(* CODESYS project liang test485.project

Project tree, tasks and I/O mapping:
  Device : AM402-CPU1608TP/TN, Shenzhen Inovance Control Technology, version 3.5.11.11
    application Application
      libraries: Standard, * (System)
      task MainTask (cyclic, interval 4 ms, priority 1) calls PLC_PRG
      program PLC_PRG [ST]
      DifferentialMonitor
      data type ST_MBTask
      program FB_ModbusRTU_Poller [ST]
    HardWare Configuration
    Network Configuration
      LocalBus Config
    Device Diagnosis
    Resources List
    ConfigStorage
    SoftMotion General Axis Pool
    HIGH_SPEED_IO : 高速IO模块, Inovance, version 00.00.00.20
        unmapped channels: InputData, OutputData
      HSIO
    MODBUS_COM0 : Modbus主站, inovance, version 00.00.00.10
        settings: Vendor.parameterset.Bit0 = False; Vendor.res = 0;  = 0
      modbus_protocol : Modbus Slave, Inovance, version 00.00.00.10
          settings: UseDec = False; modbus slave com port.ChannelNum = 3; modbus slave com port.EnableSlaveVariable = 1001; channel.PremeterSet.Bit2 = TRUE; channel.PremeterSet.Bit4 = TRUE; channel.CycleTimes = 500; channel.ReadRegOffSet = 0; channel.WriteRegOffSet = 8193; channel.IOChannel = 0; channel.ResendCount = 1; channel.ChannelName = '写频率'; channel.ChannelNote = ''; channel.PremeterSet.Bit2 = TRUE; channel.PremeterSet.Bit4 = TRUE; channel.ReadRegOffSet = 0; channel.WriteRegOffSet = 8192; channel.ResendCount = 1; channel.ChannelName = '写控制字'; channel.ChannelNote = ''; channel.PremeterSet.Bit3 = TRUE; channel.ReadRegOffSet = 8448; channel.ReadRegLeg = 4; channel.WriteRegOffSet = 0; channel.IOChannel = 2; channel.ResendCount = 1; channel.ChannelName = '读状态'; channel.ChannelNote = ''
          input  Application.PLC_PRG.Feedback1 AT %IW1 :  ARRAY[0..3] OF WORD  // 读状态
          output Application.PLC_PRG.Freq1 : WORD  // 写频率.写频率
          output Application.PLC_PRG.Ctrl1 :  ARRAY[0..0] OF WORD  // 写控制字
          unmapped channels: %QW1 写频率
    HwConfiguratioinDevice : SystemConfig, Inovance, version 00.00.00.10
  SMElement/
    SM0_SM511
    SM512_SM1023
    SM1024_SM1535
    SM1536_SM2047
    SM2048_SM2559
    SM2560_SM3071
    SM3072_SM3583
    SM3584_SM4095
    SM4096_SM4607
    SM4608_SM5119
    SM5120_SM5631
    SM5632_SM6143
    SM6144_SM6655
    SM6656_SM7167
    SM7168_SM7679
    SM7680_SM8191
    SM8192_SM8703
    SM8704_SM9215
    SM9216_SM9727
    SM9728_SM9999
  SDElement/
    SD0_SD511
    SD512_SD1023
    SD1024_SD1535
    SD1536_SD2047
    SD2048_SD2559
    SD2560_SD3071
    SD3072_SD3583
    SD3584_SD4095
    SD4096_SD4607
    SD4608_SD5119
    SD5120_SD5631
    SD5632_SD6143
    SD6144_SD6655
    SD6656_SD7167
    SD7168_SD7679
    SD7680_SD8191
    SD8192_SD8703
    SD8704_SD9215
    SD9216_SD9727
    SD9728_SD9999
*)

// Device/Application/ST_MBTask
TYPE ST_MBTask :
STRUCT
	 Enable : BOOL;
	 Slave: UINT;
	 FunctionCode:UINT;  //功能码3、4、6、16，十进制
	 Address:UINT;       //原始零起始寄存器偏移，不加40001
	 Quantity:WORD;
	 Data:ARRAY[0..19] OF WORD;
	 LastOK: BOOL;
	 Status:WORD;
	 LastValue0:WORD;
END_STRUCT
END_TYPE

// Device/Application/PLC_PRG
PROGRAM PLC_PRG
VAR
	Tasks:ARRAY[1..32] OF ST_MBTask;
	Bus : FB_ModbusRTU_Poller;
	RunPolling:BOOL;
	Enable1:BOOL;
	Enable2:BOOL;
	Enable3:BOOL;
	Ctrl1:WORD;
	Ctrl2:WORD;
	Ctrl3:WORD;
	Freq1:WORD;
	Freq2:WORD;
	Freq3:WORD;
	Feedback1 : ARRAY[0..3] OF WORD;
    Feedback2 : ARRAY[0..3] OF WORD;
    Feedback3 : ARRAY[0..3] OF WORD;
	ReadOK1:BOOL;
	ReadOK2:BOOL;
	ReadOK3:BOOL;
	FeedbackVail1:BOOL;
	FeedbackVail2:BOOL;
	FeedbackVail3:BOOL;
	Stale1:TON;
	Stale2:TON;
	Stale3:TON;
	DataNo:INT;
END_VAR

Tasks[1].Enable:=Enable1;
Tasks[1].Slave:=1;
Tasks[1].FunctionCode:=6;
Tasks[1].Address:=16#2001;
Tasks[1].Quantity:=1;
Tasks[1].Data[0]:=Freq1;

Tasks[2].Enable:=Enable1;
Tasks[2].Slave:=1;
Tasks[2].FunctionCode:=6;
Tasks[2].Address:=16#2000;
Tasks[2].Quantity:=1;
Tasks[2].Data[0]:=Ctrl1;

Tasks[3].Enable:=Enable1;
Tasks[3].Slave:=1;
Tasks[3].FunctionCode:=3;
Tasks[3].Address:=16#2100;
Tasks[3].Quantity:=4;

// 任务4：站号2，写频率
Tasks[4].Enable := Enable2;
Tasks[4].Slave := 2;
Tasks[4].FunctionCode := 6;
Tasks[4].Address := 16#2001;
Tasks[4].Quantity := 1;
Tasks[4].Data[0] := Freq2;

// 任务5：站号2，写控制字
Tasks[5].Enable := Enable2;
Tasks[5].Slave := 2;
Tasks[5].FunctionCode := 6;
Tasks[5].Address := 16#2000;
Tasks[5].Quantity := 1;
Tasks[5].Data[0] := Ctrl2;

// 任务6：站号2，读状态
Tasks[6].Enable := Enable2;
Tasks[6].Slave := 2;
Tasks[6].FunctionCode := 3;
Tasks[6].Address := 16#2100;
Tasks[6].Quantity := 4;


// 任务4：站号2，写频率
Tasks[7].Enable := Enable3;
Tasks[7].Slave := 3;
Tasks[7].FunctionCode := 6;
Tasks[7].Address := 16#2001;
Tasks[7].Quantity := 1;
Tasks[7].Data[0] := Freq3;

// 任务5：站号2，写控制字
Tasks[8].Enable := Enable3;
Tasks[8].Slave := 3;
Tasks[8].FunctionCode := 6;
Tasks[8].Address := 16#2000;
Tasks[8].Quantity := 1;
Tasks[8].Data[0] := Ctrl3;

// 任务6：站号2，读状态
Tasks[9].Enable := Enable3;
Tasks[9].Slave := 3;
Tasks[9].FunctionCode := 3;
Tasks[9].Address := 16#2100;
Tasks[9].Quantity := 4;

//Bus(Enable:=RunPolling,TaskCount:=9,PollDelay:=T#30MS,WatchDog:=T#10S,
//	PortError:=SD8500,Tasks:=Tasks
//	);

ReadOK1:=Tasks[3].LastOK;
ReadOK2:=Tasks[6].LastOK;
ReadOK3:=Tasks[9].LastOK;
Stale1(IN:=NOT(Bus.Completed AND (Bus.CurrentTask=3) AND ReadOK1),PT:=T#5S);
FeedbackVail1:=RunPolling AND Enable1 AND ReadOK1 AND NOT Stale1.Q AND NOT Bus.Fault;
IF Bus.Completed AND (Bus.CurrentTask=3) AND ReadOK1 THEN
	FOR DataNo:=0 TO 3 DO
		Feedback1[DataNo]:=Tasks[3].Data[DataNo];
	END_FOR;
END_IF

END_PROGRAM

// Device/Application/FB_ModbusRTU_Poller
PROGRAM FB_ModbusRTU_Poller
VAR_INPUT
	Enable:BOOL;
	TaskCount:INT;
	PollDelay:TIME;
	WatchDog:TIME;
	PortError:WORD;
END_VAR
VAR_OUTPUT
	CurrentTask:INT;
	Completed:BOOL;
	Busy:BOOL;
	Fault:BOOL;
	CoreStatus:WORD;
END_VAR
VAR_IN_OUT
	Tasks:ARRAY[1..32] OF ST_MBTask;
END_VAR
VAR

	PollState:INT;
	Index:WORD;
	Count:WORD;
	Active:ST_MBTask;
	Work:ARRAY[0..19] OF WORD;
	Flags:ARRAY[0..2] OF BOOL;
	CountArg:WORD;
	EnOut:BOOL;
	Gap:TON;
	Guard:TON;
	ScanNo:INT;
	DataNo:INT;
	Valid:BOOL;
	EndAddress:DWORD;
END_VAR

Completed:=FALSE;
Gap(IN:=(PollState=40),PT:=PollDelay);
Guard(IN:=(PollState=30),PT:=WatchDog);

// 始终执行这同一处指令。参数采用快照，等待期间不可修改。
// 功能码06的s4必须是0，不能照搬读/多寄存器写的数量！
//EnOut := ADPRW(PollState = 30, Active.Slave, Active.FunctionCode,
//               Active.Address, CountArg, Work[0], Flags);

CASE PollState OF
	0:
	IF (TaskCount>=1) AND(TaskCount<=32) THEN
		Count:=TaskCount;
		FOR ScanNo:=1 TO Count  DO
			Tasks[ScanNo].LastOK:=FALSE;
			Tasks[ScanNo].Status:=0;
		END_FOR;
		Index:=1;
		CoreStatus:=0;
		PollState:=20;
	ELSE
	    CoreStatus:=16#F002;	
	END_IF;
	20:
	IF Enable THEN
		FOR ScanNo:=1 TO Count DO
			IF Tasks[Index].Enable THEN
				Active:=Tasks[Index];
				Valid:=
				(Active.Slave>=1)AND(Active.Slave<=247)
				AND(Active.Quantity >=1);
				IF Active.FunctionCode=6 THEN
					Valid:=Valid AND (Active.Quantity=1);
				END_IF
				EndAddress:=WORD_TO_DWORD(Active.Address)+WORD_TO_DWORD(Active.Quantity);
				Valid:=Valid AND (EndAddress<65536);
				IF Valid THEN
					FOR DataNo:=0 TO 19  DO
						Work[DataNo]:=Active.Data[DataNo];
					END_FOR;
					Flags[0]:=FALSE;Flags[1]:=FALSE;Flags[2]:=FALSE;
					CountArg:=Active.Quantity;
					IF Active.FunctionCode=6 THEN
						CountArg:=0;
					END_IF
					CurrentTask:=Index;
					PollState:=30;
					EXIT;
				END_IF
				Tasks[Index].LastOK:=FALSE;
				Tasks[Index].Status:=16#F001;
			ELSE
				Tasks[Index].LastOK:=FALSE;
				Tasks[Index].Status:=0;
			END_IF
			Index:=Index+1;
			IF Index>Count THEN Index:=1;END_IF;
		END_FOR
	END_IF
	30:
	IF Flags[1] OR Flags[2] THEN
		Tasks[Index].LastOK:=Flags[1] AND NOT Flags[2];
		Tasks[Index].Status:=0;
		IF Tasks[Index].LastOK THEN
			Tasks[Index].LastValue0:=Work[0];
			IF(Active.FunctionCode=3)OR(Active.FunctionCode=4) THEN
				FOR DataNo:=0 TO WORD_TO_INT(Active.Quantity)-1 DO
					Tasks[Index].Data[DataNo]:=Work[DataNo];
				END_FOR
            END_IF
		ELSE
			Tasks[Index].Status:=PortError;
			IF PortError=0 THEN
				Tasks[Index].Status:=16#F004;
			END_IF
		END_IF
		Completed:=TRUE;
		PollState:=40;
	ELSIF Guard.Q THEN
	    Tasks[Index].LastOK:=FALSE;
		Tasks[Index].Status:=16#F003;
		CoreStatus:=16#F003;
		Fault:=TRUE;
		Completed:=TRUE;
		PollState:=90;
    END_IF
	40:
	IF Gap.Q THEN
		Index:=Index+1;
		IF Index>Count THEN
			Index:=1;
		END_IF
		PollState:=20;
	END_IF
	90:
	Fault:=TRUE;
END_CASE
Busy:=PollState=30;

END_PROGRAM
